(* IEC 61131-3 sources: RootPLC/crates/rootplc-driver/assets/examples, 11 files *)

(* ---- array-loop.st ---- *)
(* title: Arrays and FOR loops
   tags: array, FOR, loop, sum, average, index
   description: Sum and average an array with a FOR loop; indices stay inside the declared bounds. *)
FUNCTION EX_Average : REAL
VAR_INPUT
    samples : ARRAY[1..5] OF REAL;
END_VAR
VAR
    i : INT;
    total : REAL;
END_VAR
total := 0.0;
FOR i := 1 TO 5 DO
    total := total + samples[i];
END_FOR;
EX_Average := total / 5.0;
END_FUNCTION

TEST ex_average_of_five
VAR s : ARRAY[1..5] OF REAL := [1.0, 2.0, 3.0, 4.0, 5.0]; END_VAR
ASSERT_TRUE(ABS(EX_Average(s) - 3.0) < 0.001);
END_TEST

(* ---- limit-and-scale.st ---- *)
(* title: Limit, scale and convert numbers safely
   tags: LIMIT, conversion, scaling, INT_TO_REAL, REAL_TO_INT, clamp
   description: Clamp a value with LIMIT and convert between INT and REAL explicitly, as strict IEC 61131-3 requires (no implicit narrowing). *)
FUNCTION EX_PercentToRaw : INT
VAR_INPUT
    percent : REAL;
END_VAR
EX_PercentToRaw := REAL_TO_INT(LIMIT(0.0, percent, 100.0) * 100.0);
END_FUNCTION

TEST ex_percent_to_raw
ASSERT_EQ(5000, EX_PercentToRaw(50.0));
ASSERT_EQ(10000, EX_PercentToRaw(150.0));
ASSERT_EQ(0, EX_PercentToRaw(-3.0));
END_TEST

(* ---- interlock-permissive.st ---- *)
(* title: Interlock: permissives and trips
   tags: interlock, safety, permissive, trip, emergency stop, guard
   description: A drive may start only when all permissives are true; any trip stops it at once and it needs a new start. The common safety-interlock pattern. *)
FUNCTION_BLOCK EX_Interlock
VAR_INPUT
    start, stop : BOOL;
    permissive_ok, trip : BOOL;
END_VAR
VAR_OUTPUT
    run : BOOL;
END_VAR
IF stop OR trip OR NOT permissive_ok THEN
    run := FALSE;
ELSIF start THEN
    run := TRUE;
END_IF;
END_FUNCTION_BLOCK

TEST ex_trip_wins
VAR uut : EX_Interlock; END_VAR
uut(start := TRUE, permissive_ok := TRUE);
ASSERT_TRUE(uut.run);
uut(start := TRUE, trip := TRUE);
ASSERT_FALSE(uut.run);
uut(start := FALSE, trip := FALSE);
ASSERT_FALSE(uut.run);
END_TEST

(* ---- state-machine.st ---- *)
(* title: State machine with an enumeration and CASE
   tags: state machine, sequence, CASE, enum, step
   description: A three-step sequence (idle, running, done) written as an enumeration and a CASE statement; the pattern for any step sequence. *)
TYPE E_Step : (Idle, Running, Done); END_TYPE

FUNCTION_BLOCK EX_Sequence
VAR_INPUT
    go, finished, ack : BOOL;
END_VAR
VAR_OUTPUT
    state : E_Step;
    busy : BOOL;
END_VAR
CASE state OF
    E_Step#Idle:
        IF go THEN state := E_Step#Running; END_IF;
    E_Step#Running:
        IF finished THEN state := E_Step#Done; END_IF;
    E_Step#Done:
        IF ack THEN state := E_Step#Idle; END_IF;
END_CASE;
busy := state = E_Step#Running;
END_FUNCTION_BLOCK

TEST ex_sequence_steps
VAR uut : EX_Sequence; END_VAR
uut(go := TRUE);
ASSERT_TRUE(uut.busy);
uut(go := FALSE, finished := TRUE);
ASSERT_TRUE(uut.state = E_Step#Done);
uut(finished := FALSE, ack := TRUE);
ASSERT_TRUE(uut.state = E_Step#Idle);
END_TEST

(* ---- struct-record.st ---- *)
(* title: Structures as records
   tags: struct, record, data type, TYPE
   description: Group related values in a STRUCT type and pass it to a function block. *)
TYPE ST_Recipe : STRUCT
    temperature : REAL;
    duration : TIME;
    label : STRING[20];
END_STRUCT; END_TYPE

FUNCTION_BLOCK EX_Oven
VAR_INPUT
    recipe : ST_Recipe;
END_VAR
VAR_OUTPUT
    setpoint : REAL;
    hold : TIME;
END_VAR
setpoint := recipe.temperature;
hold := recipe.duration;
END_FUNCTION_BLOCK

TEST ex_recipe
VAR
    uut : EX_Oven;
    r : ST_Recipe := (temperature := 180.0, duration := T#20m, label := 'bread');
END_VAR
uut(recipe := r);
ASSERT_TRUE(ABS(uut.setpoint - 180.0) < 0.001);
ASSERT_TRUE(uut.hold = T#20m);
END_TEST

(* ---- testing-pattern.st ---- *)
(* title: How to write TEST blocks with virtual time
   tags: test, TEST, ASSERT, ADVANCE, virtual time, white-box
   description: The testing pattern: instantiate the program or block, call it once per cycle, move virtual time with ADVANCE, and assert on inputs, outputs or internal variables. *)
FUNCTION_BLOCK EX_Toggle
VAR_INPUT
    enable : BOOL;
END_VAR
VAR_OUTPUT
    lamp : BOOL;
END_VAR
VAR
    t : TON;
END_VAR
t(IN := enable AND NOT t.Q, PT := T#500ms);
IF t.Q THEN
    lamp := NOT lamp;
END_IF;
IF NOT enable THEN
    lamp := FALSE;
END_IF;
END_FUNCTION_BLOCK

TEST ex_toggle_after_half_second
VAR uut : EX_Toggle; i : INT; END_VAR
FOR i := 1 TO 6 DO uut(enable := TRUE); ADVANCE(T#100ms); END_FOR;
ASSERT_TRUE(uut.lamp);
uut(enable := FALSE);
ASSERT_FALSE(uut.lamp);
END_TEST

(* ---- counter-preset.st ---- *)
(* title: Up-counter with preset and reset
   tags: counter, CTU, count, preset, batch
   description: Count parts with CTU until a preset is reached; reset starts a new batch. *)
PROGRAM EX_Batch
VAR_INPUT
    part, reset : BOOL;
END_VAR
VAR_OUTPUT
    batch_full : BOOL;
    count : INT;
END_VAR
VAR
    c : CTU;
END_VAR
c(CU := part, R := reset, PV := 5);
batch_full := c.Q;
count := c.CV;
END_PROGRAM

TEST ex_batch_of_five
VAR uut : EX_Batch; i : INT; END_VAR
FOR i := 1 TO 5 DO uut(part := TRUE); uut(part := FALSE); END_FOR;
ASSERT_TRUE(uut.batch_full);
ASSERT_EQ(5, uut.count);
uut(reset := TRUE);
ASSERT_EQ(0, uut.count);
END_TEST

(* ---- edge-detect.st ---- *)
(* title: Rising and falling edge detection
   tags: edge, R_TRIG, F_TRIG, pulse, one-shot, button
   description: Detect a rising and a falling edge of a signal with the standard blocks R_TRIG and F_TRIG; the outputs are TRUE for one cycle. *)
PROGRAM EX_EdgeDetect
VAR_INPUT
    button : BOOL;
END_VAR
VAR_OUTPUT
    pressed, released : BOOL;
END_VAR
VAR
    up : R_TRIG;
    down : F_TRIG;
END_VAR
up(CLK := button);
down(CLK := button);
pressed := up.Q;
released := down.Q;
END_PROGRAM

TEST ex_edge_one_cycle
VAR uut : EX_EdgeDetect; END_VAR
uut(button := TRUE);
ASSERT_TRUE(uut.pressed);
uut(button := TRUE);
ASSERT_FALSE(uut.pressed);
uut(button := FALSE);
ASSERT_TRUE(uut.released);
END_TEST

(* ---- flip-flops.st ---- *)
(* title: Set and reset flip-flops (SR, RS)
   tags: SR, RS, flip-flop, latch, set, reset, priority
   description: SR gives set priority, RS gives reset priority; choose RS when the reset is a safety condition. *)
PROGRAM EX_FlipFlops
VAR_INPUT
    s, r : BOOL;
END_VAR
VAR_OUTPUT
    set_wins, reset_wins : BOOL;
END_VAR
VAR
    a : SR;
    b : RS;
END_VAR
a(S1 := s, R := r);
b(S := s, R1 := r);
set_wins := a.Q1;
reset_wins := b.Q1;
END_PROGRAM

TEST ex_priorities
VAR uut : EX_FlipFlops; END_VAR
uut(s := TRUE, r := TRUE);
ASSERT_TRUE(uut.set_wins);
ASSERT_FALSE(uut.reset_wins);
END_TEST

(* ---- motion-shuttle.st ---- *)
(* title: Motion: shuttle between two positions on one axis
   tags: motion, axis, servo, MC_Power, MC_Home, MC_MoveAbsolute, RootMotion, PLCopen
   description: A shuttle axis powers up, homes, then moves to a load or unload position with MC_MoveAbsolute (trapezoid profile). The virtual axis lets the TEST check timing, speed and the final position before a real drive is connected.
   libraries: RootMotion *)
PROGRAM EX_Shuttle
VAR_INPUT
    run        : BOOL;     (* power the shuttle *)
    goUnload   : BOOL;     (* TRUE: unload position, FALSE: load position *)
END_VAR
VAR_OUTPUT
    atLoad, atUnload : BOOL;
    failed           : BOOL;
END_VAR
VAR
    shuttle  : AXIS_REF;   (* mm *)
    enableAx : MC_Power;
    reference : MC_Home;
    toLoad   : MC_MoveAbsolute;
    toUnload : MC_MoveAbsolute;
END_VAR
shuttle.CycleTime := 0.01; (* this program runs every 10 ms *)
enableAx(Enable := run, Axis := shuttle);
reference(Execute := enableAx.Status, Position := 0.0, Axis := shuttle);
toUnload(Execute := run AND shuttle.Homed AND goUnload, Position := 500.0,
         Velocity := 250.0, Acceleration := 1000.0, Deceleration := 1000.0, Axis := shuttle);
toLoad(Execute := run AND shuttle.Homed AND NOT goUnload, Position := 0.0,
       Velocity := 250.0, Acceleration := 1000.0, Deceleration := 1000.0, Axis := shuttle);
RP_VirtualAxis(Axis := shuttle);
atUnload := toUnload.Done;
atLoad := shuttle.Homed AND NOT goUnload AND shuttle.State = MC_AXIS_STATE#Standstill
          AND ABS(shuttle.Position) < 0.001;
failed := enableAx.Error; (* the axis is in ErrorStop, e.g. after a software limit *)
END_PROGRAM

TEST ex_shuttle_unload_and_back
VAR uut : EX_Shuttle; i : INT; arrived : INT := -1; END_VAR
uut(run := TRUE);
uut(run := TRUE);
ASSERT_TRUE(uut.atLoad);
FOR i := 1 TO 300 DO
    uut(run := TRUE, goUnload := TRUE);
    ASSERT_TRUE(uut.shuttle.Velocity <= 250.0001);
    IF uut.atUnload AND arrived < 0 THEN arrived := i; END_IF;
END_FOR;
(* 0.25 s up + 1.75 s cruise + 0.25 s down = 2.25 s, Done one cycle later *)
ASSERT_TRUE(arrived >= 225 AND arrived <= 228);
ASSERT_TRUE(ABS(uut.shuttle.Position - 500.0) < 0.000001);
FOR i := 1 TO 300 DO uut(run := TRUE, goUnload := FALSE); END_FOR;
ASSERT_TRUE(uut.atLoad);
ASSERT_FALSE(uut.failed);
END_TEST

TEST ex_shuttle_off_stops_the_axis
VAR uut : EX_Shuttle; i : INT; END_VAR
uut(run := TRUE);
FOR i := 1 TO 50 DO uut(run := TRUE, goUnload := TRUE); END_FOR;
uut(run := FALSE, goUnload := TRUE);
ASSERT_TRUE(uut.shuttle.State = MC_AXIS_STATE#Disabled);
ASSERT_TRUE(uut.shuttle.Velocity = 0.0);
ASSERT_FALSE(uut.atUnload);
END_TEST

TEST ex_shuttle_flags_only_when_true
VAR uut : EX_Shuttle; i : INT; END_VAR
FOR i := 1 TO 5 DO uut(run := FALSE); END_FOR;
ASSERT_FALSE(uut.atLoad);
ASSERT_FALSE(uut.failed);
uut(run := TRUE);
FOR i := 1 TO 20 DO uut(run := TRUE, goUnload := TRUE); END_FOR;
ASSERT_FALSE(uut.atLoad);
ASSERT_FALSE(uut.atUnload);
(* a software limit before the unload position stops the axis with an error *)
uut.shuttle.LimitsEnabled := TRUE;
uut.shuttle.PositiveLimit := 400.0;
uut.shuttle.NegativeLimit := -10.0;
FOR i := 1 TO 300 DO uut(run := TRUE, goUnload := TRUE); END_FOR;
ASSERT_TRUE(uut.failed);
ASSERT_FALSE(uut.atUnload);
ASSERT_TRUE(uut.shuttle.Position <= 400.0);
FOR i := 1 TO 300 DO uut(run := TRUE, goUnload := FALSE); END_FOR;
ASSERT_FALSE(uut.atLoad);
END_TEST

(* ---- on-off-delay.st ---- *)
(* title: On-delay and off-delay timers
   tags: timer, TON, TOF, delay, time
   description: Switch an output on 2 s after a request and keep a fan running 5 s after the request ends, with TON and TOF. *)
PROGRAM EX_Delays
VAR_INPUT
    request : BOOL;
END_VAR
VAR_OUTPUT
    heater_on, fan_on : BOOL;
END_VAR
VAR
    on_delay : TON;
    run_on : TOF;
END_VAR
on_delay(IN := request, PT := T#2s);
run_on(IN := request, PT := T#5s);
heater_on := on_delay.Q;
fan_on := run_on.Q;
END_PROGRAM

TEST ex_delays_on_and_run_on
VAR uut : EX_Delays; i : INT; END_VAR
FOR i := 1 TO 15 DO uut(request := TRUE); ADVANCE(T#100ms); END_FOR;
ASSERT_FALSE(uut.heater_on);
FOR i := 1 TO 10 DO uut(request := TRUE); ADVANCE(T#100ms); END_FOR;
uut(request := TRUE);
ASSERT_TRUE(uut.heater_on);
FOR i := 1 TO 30 DO uut(request := FALSE); ADVANCE(T#100ms); END_FOR;
ASSERT_TRUE(uut.fan_on);
FOR i := 1 TO 30 DO uut(request := FALSE); ADVANCE(T#100ms); END_FOR;
ASSERT_FALSE(uut.fan_on);
END_TEST
